{attribute 'linkalways'}
{attribute 'no_explicit_call' := 'Use the methods of this class'}
{attribute 'enable_dynamic_creation'}
FUNCTION_BLOCK SweepMission
VAR
	_state : MissionState := MissionState.IDLE;
	stateBeforePause : MissionState;
	lastSequence : UDINT;
	_desiredTwist : Twist;
	_hasMap : BOOL;
	requestedPose : Pose2D;
	hasPoseRequest : BOOL;
	hasMapClearRequest : BOOL;
END_VAR

METHOD Execute
IF RobotHmi.command.sequence <> lastSequence THEN
	lastSequence := RobotHmi.command.sequence;
	Handle(RobotHmi.command.code);
	RobotHmi.status.acknowledgedSequence := lastSequence;
END_IF

CASE _state OF
	MissionState.MANUAL:
		_desiredTwist := RobotHmi.command.manualTwist;
	MissionState.MAPPING:
		// Til roboten kan utforske selv (M5), kjører du den med tastaturet mens den kartlegger.
		_desiredTwist := RobotHmi.command.manualTwist;
	MissionState.SWEEPING, MissionState.RETURNING_TO_DOCK:
		// Kommer i M6: feiing og retur til lader.
		_desiredTwist := Stopped();
ELSE
	_desiredTwist := Stopped();
END_CASE

RobotHmi.status.missionState := _state;
RobotHmi.status.hasMap := _hasMap;
END_METHOD

METHOD PRIVATE Handle
VAR_INPUT
	code : HmiCommandCode;
END_VAR
RobotHmi.status.lastRejection := '';

IF code = HmiCommandCode.EMERGENCY_STOP THEN
	_state := MissionState.EMERGENCY_STOPPED;
	RETURN;
END_IF
IF code = HmiCommandCode.SET_POSE THEN
	IF IsBusy() THEN
		Reject('Stopp oppdraget før du setter posisjonen.');
	ELSE
		requestedPose := RobotHmi.command.pose;
		hasPoseRequest := TRUE;
	END_IF
	RETURN;
END_IF
IF _state = MissionState.EMERGENCY_STOPPED AND code <> HmiCommandCode.RESET THEN
	Reject('Nødstopp er aktiv. Tilbakestill først.');
	RETURN;
END_IF

CASE code OF
	HmiCommandCode.RESET:
		_state := MissionState.IDLE;
	HmiCommandCode.MANUAL_DRIVE:
		IF IsBusy() THEN
			Reject('Stopp oppdraget før du kjører manuelt.');
		ELSE
			_state := MissionState.MANUAL;
		END_IF
	HmiCommandCode.START_MAPPING:
		// Et nytt kart hver gang. Fortsetter du etter en pause, bruker du RESUME.
		_state := MissionState.MAPPING;
		_hasMap := FALSE;
		hasMapClearRequest := TRUE;
	HmiCommandCode.START_SWEEPING:
		IF _hasMap THEN
			_state := MissionState.SWEEPING;
		ELSE
			Reject('Kartet mangler. Kjør kartlegging først.');
		END_IF
	HmiCommandCode.PAUSE:
		IF IsBusy() THEN
			stateBeforePause := _state;
			_state := MissionState.PAUSED;
		ELSE
			Reject('Det er ikke noe oppdrag å pause.');
		END_IF
	HmiCommandCode.RESUME:
		IF _state = MissionState.PAUSED THEN
			_state := stateBeforePause;
		ELSE
			Reject('Det er ikke noe pauset oppdrag.');
		END_IF
	HmiCommandCode.STOP:
		IF _state = MissionState.MAPPING OR (_state = MissionState.PAUSED AND stateBeforePause = MissionState.MAPPING) THEN
			_hasMap := TRUE;
		END_IF
		_state := MissionState.IDLE;
	HmiCommandCode.GO_TO_DOCK:
		_state := MissionState.RETURNING_TO_DOCK;
END_CASE
END_METHOD

METHOD PRIVATE IsBusy : BOOL
IsBusy := _state = MissionState.MAPPING OR _state = MissionState.SWEEPING OR _state = MissionState.RETURNING_TO_DOCK;
END_METHOD

METHOD PRIVATE Reject
VAR_INPUT
	reason : STRING(80);
END_VAR
RobotHmi.status.lastRejection := reason;
END_METHOD

METHOD PRIVATE Stopped : Twist
VAR
	standingStill : Twist;
END_VAR
Stopped := standingStill;
END_METHOD

METHOD TryTakePoseRequest : BOOL
VAR_INPUT
	pose : REFERENCE TO Pose2D;
END_VAR
IF NOT hasPoseRequest THEN
	RETURN;
END_IF
pose := requestedPose;
hasPoseRequest := FALSE;
TryTakePoseRequest := TRUE;
END_METHOD

// TRUE én gang når en ny kartlegging starter, så kartet kan tømmes.
METHOD TryTakeMapClearRequest : BOOL
TryTakeMapClearRequest := hasMapClearRequest;
hasMapClearRequest := FALSE;
END_METHOD

PROPERTY State : MissionState
GET
State := _state;
END_GET
END_PROPERTY

PROPERTY DesiredTwist : Twist
GET
DesiredTwist := _desiredTwist;
END_GET
END_PROPERTY

PROPERTY ShouldDrive : BOOL
GET
ShouldDrive := _state = MissionState.MANUAL OR IsBusy();
END_GET
END_PROPERTY

END_FUNCTION_BLOCK

(* stored: Version 1.1.0.1, ProductVersion 3.1.4026.12
   POU SweepMission: Id {e41591d1-bb67-5c93-93c1-653c454fd246}, SpecialFunc None
   Method Execute: Id {0edb486b-e6d2-5352-ac1f-a2f72835a724}
   Method Handle: Id {b572e568-37ab-508b-b7c6-42fbd5147f7e}
   Method IsBusy: Id {eda4ea94-5c3e-599c-aad6-57368444694f}
   Method Reject: Id {29783acd-ce63-5b0b-b23a-8706aa79491f}
   Method Stopped: Id {79198e0b-a880-5d10-9263-47f1f8f4786f}
   Method TryTakePoseRequest: Id {306f9d1e-d706-40a5-91e6-e021f48d4ace}
   Method TryTakeMapClearRequest: Id {1fb4962b-93da-42cd-95fe-e8c20436d1bb}
   Property State: Id {dbdbf95e-8f4b-5a68-9ddb-a6be58b8826a}
   Get Get: Id {bb6bc095-2963-5642-bdbb-9e67613a7d7e}
   Property DesiredTwist: Id {b9558c05-0211-5579-82fb-906b1dff166c}
   Get Get: Id {a3c88e9d-a866-53f0-a45a-d5c638ad65c5}
   Property ShouldDrive: Id {148580db-2e22-5441-b6bc-6a52e4c70a85}
   Get Get: Id {34c545f2-47da-5fc5-b10b-7f2406f59224} *)
